FUNCTION_BLOCK FB_PI_Controller (* Migrated from IEC 61131-3 ST *)
  (* Standard: 61499-2 *)
  (* Version 1.0, 2026-11-06, st2fb *)
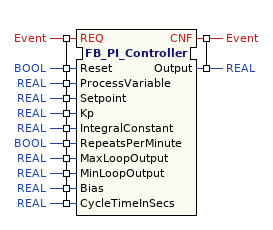
  EVENT_INPUT
    REQ WITH Reset, ProcessVariable, Setpoint, Kp, IntegralConstant, RepeatsPerMinute, MaxLoopOutput, MinLoopOutput, Bias, CycleTimeInSecs;
  END_EVENT
  EVENT_OUTPUT
    CNF WITH Output;
  END_EVENT
  VAR_INPUT
    Reset : BOOL;
    ProcessVariable : REAL;
    Setpoint : REAL;
    Kp : REAL;
    IntegralConstant : REAL;
    RepeatsPerMinute : BOOL := TRUE;
    MaxLoopOutput : REAL;
    MinLoopOutput : REAL;
    Bias : REAL;
    CycleTimeInSecs : REAL;
  END_VAR
  VAR_OUTPUT
    Output : REAL;
  END_VAR
  VAR
    preClampedOutput : REAL;
    p_Term : REAL;
    i_Term : REAL;
    i_Ki : REAL;
    i_Pause : BOOL;
    i_Ki2 : REAL;
    i_integral : REAL;
    i_error : REAL;
    i_Max : REAL := 1000.0;
    i_Min : REAL := -1000.0;
    i_done : BOOL;
  END_VAR
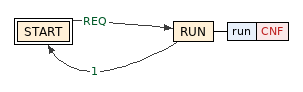
  EC_STATES
    START;
    RUN : run -> CNF;
  END_STATES
  EC_TRANSITIONS
    START TO RUN := REQ;
    RUN TO START := 1;
  END_TRANSITIONS
  ALGORITHM run IN ST:
p_Term := (Setpoint - ProcessVariable) * Kp;

i_Ki := IntegralConstant / SEL(RepeatsPerMinute, 1.0, 60.0);
i_Pause := ((preClampedOutput > MaxLoopOutput) AND (ProcessVariable < Setpoint)) OR ((preClampedOutput < MinLoopOutput) AND (ProcessVariable > Setpoint));
i_done := FALSE;
IF i_Ki <= 0.0 THEN
  i_Term := 0.0;
  i_done := TRUE;
END_IF;
IF NOT i_done THEN
  IF Reset THEN
    i_integral := 0.0;
  ELSIF i_Pause THEN
    i_done := TRUE;
  END_IF;
END_IF;
IF NOT i_done THEN
  i_Ki2 := i_Ki * CycleTimeInSecs;
  i_error := Setpoint - ProcessVariable;
  i_integral := i_integral + i_Ki2 * i_error;
  IF i_integral > i_Max THEN
    i_integral := i_Max;
  ELSIF i_integral < i_Min THEN
    i_integral := i_Min;
  END_IF;
  i_Term := i_integral;
END_IF;

preClampedOutput := p_Term + i_Term + Bias;
Output := LIMIT(MinLoopOutput, preClampedOutput, MaxLoopOutput);
  END_ALGORITHM
END_FUNCTION_BLOCK
